(* LS Electric XG5000 project: NewProject *)
(* PLC LSPLC *)
(* task ControlLoop: Kind=2 Priority=7 Device=250 *)
(* task Initialize: Kind=1 Priority=2 *)
(* task Trigger0: Kind=3 Priority=2 Device=%MX0 *)
(* task Trigger1: Kind=3 Priority=3 Device=%MX0 BitCondition=1 *)
(* task Trigger2: Kind=3 Priority=4 Device=%MX0 BitCondition=2 *)
(* task Trigger3: Kind=3 Priority=5 Device=%MX0 BitCondition=3 *)
(* task Trigger4: Kind=3 Priority=6 Device=%MX0 BitCondition=4 *)
(* task Trigger5: Kind=3 Priority=7 Device=%MW0 WordValue=65535 *)
(* task Trigger6: Kind=3 Priority=2 Device=%MW0 WordValue=65535 WordCondition=1 *)
(* task Trigger7: Kind=3 Priority=3 Device=%MW0 WordValue=65535 WordCondition=2 *)
(* task Trigger8: Kind=3 Priority=4 Device=%MW0 WordValue=65535 WordCondition=3 *)
(* task Trigger9: Kind=3 Priority=5 Device=%MW0 WordValue=65535 WordCondition=4 *)

PROGRAM ScanLoop (* task: 스캔 프로그램 *)

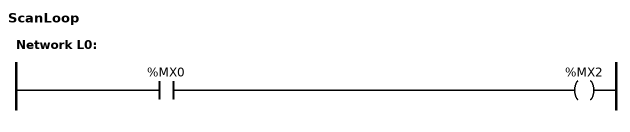
(* Rung L0 *)
%MX2 := %MX0;
END_PROGRAM

PROGRAM NewProgram (* task: ControlLoop *)

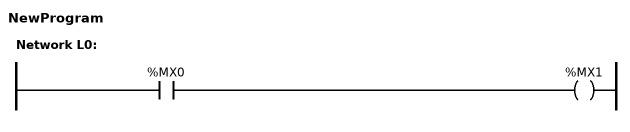
(* Rung L0 *)
%MX1 := %MX0;
END_PROGRAM

PROGRAM Worker0 (* task: Trigger0 *)

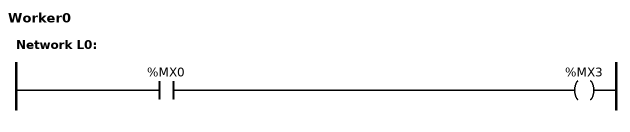
(* Rung L0 *)
%MX3 := %MX0;
END_PROGRAM

PROGRAM Worker1 (* task: Trigger1 *)

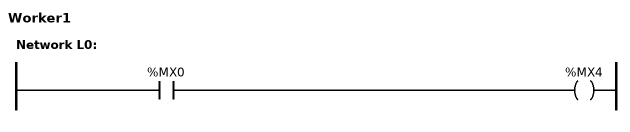
(* Rung L0 *)
%MX4 := %MX0;
END_PROGRAM

PROGRAM Worker2 (* task: Trigger2 *)

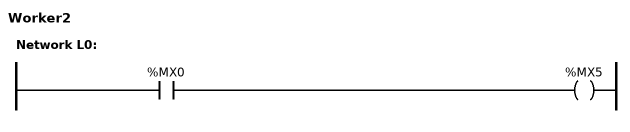
(* Rung L0 *)
%MX5 := %MX0;
END_PROGRAM

PROGRAM Worker3 (* task: Trigger3 *)

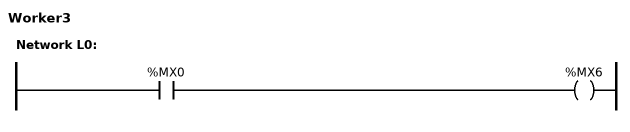
(* Rung L0 *)
%MX6 := %MX0;
END_PROGRAM

PROGRAM Worker4 (* task: Trigger4 *)

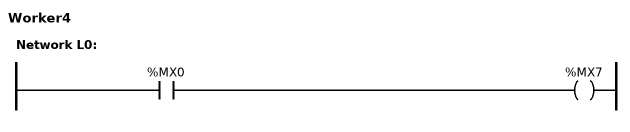
(* Rung L0 *)
%MX7 := %MX0;
END_PROGRAM

PROGRAM Worker5 (* task: Trigger5 *)

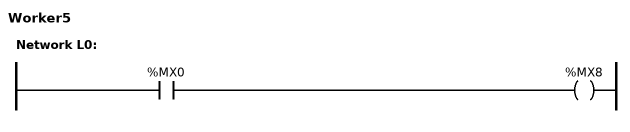
(* Rung L0 *)
%MX8 := %MX0;
END_PROGRAM

PROGRAM Worker6 (* task: Trigger6 *)

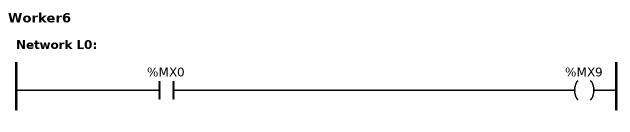
(* Rung L0 *)
%MX9 := %MX0;
END_PROGRAM

PROGRAM Worker7 (* task: Trigger7 *)

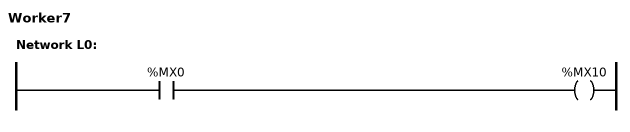
(* Rung L0 *)
%MX10 := %MX0;
END_PROGRAM

PROGRAM Worker8 (* task: Trigger8 *)

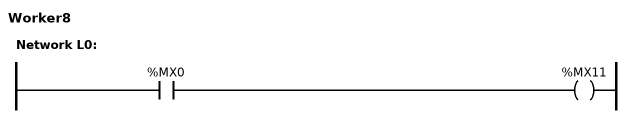
(* Rung L0 *)
%MX11 := %MX0;
END_PROGRAM

PROGRAM Worker9 (* task: Trigger9 *)

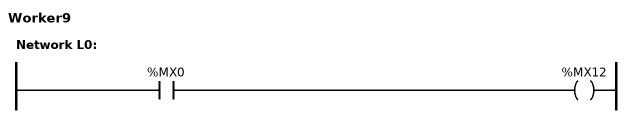
(* Rung L0 *)
%MX12 := %MX0;
END_PROGRAM